Fanuc KAREL source: KA00162.KL

PROGRAM KA00162
%NOLOCKGROUP
VAR
  SRC: ARRAY[4] OF REAL
  DST: ARRAY[4] OF JOINTPOS
BEGIN
  DST = SRC
END KA00162
